    rq_activate_all_grippers(True)
    # end: URCap Program Node
  end
  $ 62 "zero_ftsensor()"
  zero_ftsensor()
  $ 63 "EXTT"
  $ 64 "Set GRP_3F_Enable=Off"
  set_standard_digital_out(4, False)
  $ 65 "Set BarcodeTrigger=Off"
  set_standard_digital_out(6, False)
  $ 66 "Set GRP_3F_Decap=Off"
  set_standard_digital_out(3, False)
  $ 67 "Set GRP_3F_Cap=Off"
  set_standard_digital_out(2, False)
  $ 68 "Set GRP_3F_Open=Off"
  set_standard_digital_out(5, False)
  $ 69 "PSE_T≔get_tool_free_pose(dir=[0,0,0.150], move_in_base_frame=True)"
  global PSE_T=get_tool_free_pose(dir=[0,0,0.150], move_in_base_frame=True)
  $ 70 "If is_reachable(Base_const, [PSE_T])"
  if (is_reachable(p[0.0,0.0,0.0,0.0,0.0,0.0], [PSE_T])):
    $ 71 "MoveL"
    $ 72 "PSE_T" "breakAfter"
    movel(PSE_T, a=1.2, v=0.15)
  end
  $ 74 "powder dispensing variable init"
  $ 75 "Start_thread≔ False "
  global Start_thread=  False
  $ 76 "vib_thread≔ False "
  global vib_thread=  False
  $ 77 "kp≔0.0015"
  global kp=0.0015
  $ 78 "ki≔0.0001"
  global ki=0.0001
  $ 79 "kd≔0.01"
  global kd=0.01
  $ 80 "dt≔0.03"
  global dt=0.03
  $ 81 "Integral_error≔0"
  global Integral_error=0
  $ 82 "current_error≔0"
  global current_error=0
  $ 83 "previous_error≔0"
  global previous_error=0
  $ 84 "tilt_increment≔0"
  global tilt_increment=0
  $ 85 "tilt_angle≔0"
  global tilt_angle=0
  $ 86 "diff≔0"
  global diff=0
  $ 87 "current_pose≔get_actual_tcp_pose()"
  global current_pose= get_actual_tcp_pose ()
  $ 88 "Relative_trans≔p[0, 0, -0.035, 0, 0, 0]"
  global Relative_trans=p[0, 0, -0.035, 0, 0, 0]
  $ 89 "ContA_plc_offst≔p[-0.00205, 0.02547, 0.03730, -0.03, -2.183, 6.165]"
  global ContA_plc_offst=p[-0.00205, 0.02547, 0.03730, -0.03, -2.183, 6.165]
  $ 90 "PowA_50_offset≔p[0.21808, -0.19943, 0.06584, 0, 0, 0]"
  global PowA_50_offset=p[0.21808, -0.19943, 0.06584, 0, 0, 0]
  $ 92 "tilt_init_reference()"
  tilt_init_reference()
  $ 93 "switch_spat_M≔ True "
  global switch_spat_M=  True
  $ 94 "switch_spat_S≔ True "
  global switch_spat_S=  True
  $ 95 "switch_spat_F_M≔ True "
  global switch_spat_F_M=  True
  $ 96 "switch_spat_F_S≔ True "
  global switch_spat_F_S=  True
  $ 97 "last_scale≔0"
  global last_scale=0
  $ 98 "W_EMPTY≔51.381"
  global W_EMPTY=51.381
  $ 771 "Thread_1"
  thread Thread_1():
    while (True):
      $ 772 "If Start_thread≟ True "
      if (Start_thread ==   True  ):
        $ 773 "weight_value≔get_weight()"
        global weight_value=get_weight()
        $ 774 "Wait: 0.1"
        sleep(0.1)
        $ 775 "sync()"
        sync()
      end
      $ 776 "sync()"
      sync()
    end
  end
  threadId_Thread_1 = run Thread_1()
  $ 777 "Thread_2"
  thread Thread_2():
    while (True):
      $ 778 "Loop vib_thread≟ True "
      thread Thread_while_778():
        while (True):
          $ 779 "diff≔target_weight-weight_value"
          global diff=target_weight-weight_value
          $ 780 "If diff>0.02 and spatula≠'spatula_flat_S'"
          global thread_flag_780=0
          thread Thread_if_780():
            $ 782 "Set AO[0]=4.0"
            set_standard_analog_out(0, 0.4)
            thread_flag_780 = 1
          end
          if (diff>0.02  and  spatula != "spatula_flat_S"):
            global thread_handler_780=run Thread_if_780()
            while (thread_flag_780 == 0):
              if not(diff>0.02  and  spatula != "spatula_flat_S"):
                kill thread_handler_780
                thread_flag_780 = 2
              else:
                sync()
              end
            end
          else:
            thread_flag_780 = 2
          end
          if (thread_flag_780 == 2):
            $ 783 "ElseIf diff>0.02 and spatula≟'spatula_flat_S'"
            if (diff>0.02 and spatula == "spatula_flat_S"):
              $ 784 "vibration_3()"
              vibration_3()
            else:
              $ 785 "ElseIf diff≤0.03"
              global thread_flag_785=0
              thread Thread_if_785():
                $ 786 "vibration_2()"
                vibration_2()
                thread_flag_785 = 1
              end
              if (diff <= 0.03):
                global thread_handler_785=run Thread_if_785()
                while (thread_flag_785 == 0):
                  if not(diff <= 0.03):
                    kill thread_handler_785
                    thread_flag_785 = 2
                  else:
                    sync()
                  end
                end
              else:
                thread_flag_785 = 2
              end
              if (thread_flag_785 == 2):
                $ 791 "Else" "noBreak"
                $ 792 "Set AO[0]=0.0"
                set_standard_analog_out(0, 0.0)
              end
            end
          end
        end
      end
      if (vib_thread ==   True  ):
        global thread_handler_778=run Thread_while_778()
        while (vib_thread ==   True  ):
          sync()
        end
        kill thread_handler_778
      end
      $ 793 "sync()"
      sync()
    end
  end
  threadId_Thread_2 = run Thread_2()
  while (True):
    $ 99 "Robot Program"
    $ 100 "MAIN"
    $ 101 "command_manager(external_control='uGO', cond_suspend=(ITM_Manipulated and AMR_AtTarget and AMR_Charging and AMR_Battery<40), cond_unsuspend=(AMR_Battery≟60))"
    command_manager(external_control="uGO", cond_suspend=(ITM_Manipulated  and  AMR_AtTarget  and  AMR_Charging  and  AMR_Battery<40), cond_unsuspend=(AMR_Battery == 60))
    $ 102 "log_state(STATE_Info)"
    log_state(STATE_Info)
    $ 103 "Switch STATE"
    switch_1 = STATE
    $ 104 "Case 1"
    if (1 == switch_1):
      $ 105 "Stopping"
      $ 106 "STATE_Info≔'Stopping'"
      global STATE_Info="Stopping"
      $ 107 "end_freedrive_mode()"
      end_freedrive_mode()
      $ 108 "Set"
      set_tcp(p[0.0,0.0,0.161,3.1415,0.0,0.0])
      $ 109 "PSE_T≔get_tool_free_pose(dir=[0,0,0.150], move_in_base_frame=True)"
      global PSE_T=get_tool_free_pose(dir=[0,0,0.150], move_in_base_frame=True)
      $ 110 "If is_reachable(Base_const, [PSE_T])"
      if (is_reachable(p[0.0,0.0,0.0,0.0,0.0,0.0], [PSE_T])):
        $ 111 "MoveL"
        $ 112 "PSE_T" "breakAfter"
        movel(PSE_T, a=1.2, v=0.15)
      end
      $ 113 "do_transition(keep_rxry=OBJ_Picked, r=0)"
      do_transition(keep_rxry=OBJ_Picked, r=0)
      $ 122 "Call Sub_AMR_MiR_V3"
      Sub_AMR_MiR_V3()
      $ 123 "If stopping() and AMR_Done"
      if (stopping()  and  AMR_Done):
        $ 124 "STATE≔2"
        global STATE=2
        $ 125 "ugo_update_outputs()"
        ugo_update_outputs()
      end
    elif (2 == switch_1):
      $ 126 "Case 2"
      $ 127 "Stopped"
      $ 128 "STATE_Info≔'Stopped'"
      global STATE_Info="Stopped"
      $ 129 "Call Sub_AMR_MiR_V3"
      Sub_AMR_MiR_V3()
      $ 130 "If CMD_Reset  or PB_Start"
      if (CMD_Reset   or  get_standard_digital_in(0)):
        $ 131 "STATE≔3"
        global STATE=3
        $ 132 "ugo_update_outputs()"
        ugo_update_outputs()
      end
    elif (3 == switch_1):
      $ 133 "Case 3"
      $ 134 " Resetting"
      $ 135 "STATE_Info≔'Resetting'"
      global STATE_Info="Resetting"
      $ 136 "uML"
      $ 137 "reset_error()"
      reset_error()
      $ 138 "reset_warning()"
      reset_warning()
      $ 139 "PROCESS_Step≔0"
      global PROCESS_Step=0
      $ 140 "PROCESS_Info≔''"
      global PROCESS_Info=""
      $ 141 "ARM_Referenced≔ False "
      global ARM_Referenced=  False
      $ 142 "WRK_Done≔ False "
      global WRK_Done=  False
      $ 143 "ITM_Prepared≔ False "
      global ITM_Prepared=  False
      $ 144 "ITM_Manipulated≔ False "
      global ITM_Manipulated=  False
      $ 145 "STP≔0"
      global STP=0
      $ 146 "Action≔0"
      global Action=0
      $ 147 "Action_Info≔''"
      global Action_Info=""
      $ 148 "ITM_ID≔0"
      global ITM_ID=0
      $ 149 "JIG≔0"
      global JIG=0
      $ 150 "JIG_Slot≔0"
      global JIG_Slot=0
      $ 151 "Task_info≔''"
      global Task_info=""
      $ 152 "Set"
      set_tcp(p[0.0,0.0,0.161,3.1415,0.0,0.0])
      $ 153 "App"
      $ 154 "'ADD APPLICATION SPECIFIC COMMANDS'"
      # 'ADD APPLICATION SPECIFIC COMMANDS'
      $ 155 "OBJ_Type≔0"
      global OBJ_Type=0
      $ 156 "OBJ_Nbr≔0"
      global OBJ_Nbr=0
      $ 157 "If CNT_Rack_Output≥50"
      if (CNT_Rack_Output >= 50):
        $ 158 "CNT_Rack_Output≔0"
        global CNT_Rack_Output=0
      end
      $ 159 "TASK≔struct(ID=0, NAVI=struct(target=0, footprint=0, protectiveOff=0, dock=0), WORK=struct(ITM_ID_Src=0, JIG_ID_Src=0, OBJ_Nbr_Src=0, ACT_Src=0, ITM_ID_Tgt=0, JIG_ID_Tgt=0, OBJ_Nbr_Tgt=0, ACT_Tgt=0, OBJ_Type=0))"
      global TASK=struct(ID=0, NAVI=struct(target=0, footprint=0, protectiveOff=0, dock=0), WORK=struct(ITM_ID_Src=0, JIG_ID_Src=0, OBJ_Nbr_Src=0, ACT_Src=0, ITM_ID_Tgt=0, JIG_ID_Tgt=0, OBJ_Nbr_Tgt=0, ACT_Tgt=0, OBJ_Type=0))
      $ 160 "Call Sub_AMR_MiR_V3"
      Sub_AMR_MiR_V3()
      $ 161 "If resetting() and AMR_Done"
      if (resetting()  and  AMR_Done):
        $ 162 "STATE≔4"
        global STATE=4
        $ 163 "ugo_update_outputs()"
        ugo_update_outputs()
      end
    elif (4 == switch_1):
      $ 164 "Case 4"
      $ 165 "Idle"
      $ 166 "STATE_Info≔'Idle'"
      global STATE_Info="Idle"
      $ 167 "If CMD_Start"
      if (CMD_Start):
        $ 168 "STATE≔5"
        global STATE=5
        $ 169 "ugo_update_outputs()"
        ugo_update_outputs()
      end
    elif (5 == switch_1):
      $ 170 "Case 5"
      $ 171 "Starting"
      $ 172 "STATE_Info≔'Starting'"
      global STATE_Info="Starting"
      $ 173 "'ADD COMMANDS WHAT TO START WITH'"
      # 'ADD COMMANDS WHAT TO START WITH'
      $ 174 "Call Sub_AMR_MiR_V3"
      Sub_AMR_MiR_V3()
      $ 175 "get ugo data"
      $ 176 "Assign Tasks"
      $ 177 "TASK.ID = ugo_get_task()"
      TASK.ID = ugo_get_task()
      $ 178 "If TASK.ID≟1"
      if (TASK.ID == 1):
        $ 179 "Task_info≔'Charge'"
        global Task_info="Charge"
        $ 180 "Parameters"
        $ 181 "AMR_PosTarget≔1"
        global AMR_PosTarget=1
      else:
        $ 182 "ElseIf TASK.ID≟9"
        if (TASK.ID == 9):
          $ 183 "'Pick Sarstedt Rack from Variable source'"
          # 'Pick Sarstedt Rack from Variable source'
          $ 184 "Task_info≔'Navigate to Target'"
          global Task_info="Navigate to Target"
          $ 185 "Parameters"
          $ 186 "AMR_PosTarget≔UGO.read_input('00','ITM_ID')"
          global AMR_PosTarget=UGO.read_input("00","ITM_ID")
        else:
          $ 187 "ElseIf TASK.ID≟49"
          if (TASK.ID == 49):
            $ 188 "Task_info≔'Pick Containers'"
            global Task_info="Pick Containers"
            $ 189 "Parameters"
            $ 190 "ITM_ID≔1"
            global ITM_ID=1
            $ 191 "OBJ_Type≔6"
            global OBJ_Type=6
            $ 192 "JIG≔15"
            global JIG=15
            $ 193 "AMR_PosTarget≔3"
            global AMR_PosTarget=3
          else:
            $ 194 "ElseIf TASK.ID≟50"
            if (TASK.ID == 50):
              $ 195 "Task_info≔'Decap Containers'"
              global Task_info="Decap Containers"
              $ 196 "Parameters"
              $ 197 "ITM_ID≔1"
              global ITM_ID=1
              $ 198 "OBJ_Type≔6"
              global OBJ_Type=6
              $ 199 "JIG≔16"
              global JIG=16
              $ 200 "AMR_PosTarget≔5"
              global AMR_PosTarget=5
            else:
              $ 201 "ElseIf TASK.ID≟51"
              if (TASK.ID == 51):
                $ 202 "Task_info≔'Detect Spatula and transfer powder'"
                global Task_info="Detect Spatula and transfer powder"
                $ 203 "Parameters"
                $ 204 "ITM_ID≔1"
                global ITM_ID=1
                $ 205 "target_weight≔(UGO.read_input('00','Target_weight'))/1000"
                global target_weight=(UGO.read_input("00","Target_weight"))/1000
                $ 206 "OBJ_Type≔8"
                global OBJ_Type=8
                $ 207 "JIG≔16"
                global JIG=16
                $ 208 "AMR_PosTarget≔5"
                global AMR_PosTarget=5
              else:
                $ 209 "ElseIf TASK.ID≟52"
                if (TASK.ID == 52):
                  $ 210 "Task_info≔'Pick Powder'"
                  global Task_info="Pick Powder"
                  $ 211 "Parameters"
                  $ 212 "ITM_ID≔1"
                  global ITM_ID=1
                  $ 213 "OBJ_Type≔6"
                  global OBJ_Type=6
                  $ 214 "JIG≔15"
                  global JIG=15
                  $ 215 "AMR_PosTarget≔3"
                  global AMR_PosTarget=3
                else:
                  $ 216 "ElseIf TASK.ID≟53"
                  if (TASK.ID == 53):
                    $ 217 "Task_info≔'Decap Powder'"
                    global Task_info="Decap Powder"
                    $ 218 "Parameters"
                    $ 219 "ITM_ID≔1"
                    global ITM_ID=1
                    $ 220 "OBJ_Type≔6"
                    global OBJ_Type=6
                    $ 221 "JIG≔1"
                    global JIG=1
                    $ 222 "AMR_PosTarget≔5"
                    global AMR_PosTarget=5
                  else:
                    $ 223 "ElseIf TASK.ID≟54"
                    if (TASK.ID == 54):
                      $ 224 "Task_info≔'Empty and swap Powder container'"
                      global Task_info="Empty and swap Powder container"
                      $ 233 "Parameters"
                      $ 234 "ITM_ID≔1"
                      global ITM_ID=1
                      $ 236 "W_now≔(UGO.read_input('00','Container_weight'))/1000"
                      global W_now=(UGO.read_input("00","Container_weight"))/1000
                      $ 237 "Pow_name≔(UGO.read_input('00','Powder_name'))"
                      global Pow_name=(UGO.read_input("00","Powder_name"))
                      $ 238 "scooping_init()"
                      scooping_init()
                      $ 239 "target_weight≔W_now-W_EMPTY-(0.002*W_FULL)"
                      global target_weight=W_now-W_EMPTY-(0.002*W_FULL)
                      $ 240 "OBJ_Type≔6"
                      global OBJ_Type=6
                      $ 241 "JIG≔17"
                      global JIG=17
                      $ 242 "AMR_PosTarget≔5"
                      global AMR_PosTarget=5
                    else:
                      $ 243 "ElseIf TASK.ID≟55"
                      if (TASK.ID == 55):
                        $ 244 "Task_info≔'Place Powder'"
                        global Task_info="Place Powder"
                        $ 245 "Parameters"
                        $ 246 "ITM_ID≔1"
                        global ITM_ID=1
                        $ 247 "OBJ_Type≔6"
                        global OBJ_Type=6
                        $ 248 "JIG≔21"
                        global JIG=21
                        $ 249 "AMR_PosTarget≔5"
                        global AMR_PosTarget=5
                      else:
                        $ 250 "ElseIf TASK.ID≟56"
                        if (TASK.ID == 56):
                          $ 251 "Task_info≔'Dose Powder'"
                          global Task_info="Dose Powder"
                          $ 252 "Parameters"
                          $ 253 "ITM_ID≔1"
                          global ITM_ID=1
                          $ 254 "target_weight≔(UGO.read_input('00','Target_weight'))/1000"
                          global target_weight=(UGO.read_input("00","Target_weight"))/1000
                          $ 255 "W_now≔(UGO.read_input('00','Container_weight'))/1000"
                          global W_now=(UGO.read_input("00","Container_weight"))/1000
                          $ 257 "Pow_name≔(UGO.read_input('00','Powder_name'))"
                          global Pow_name=(UGO.read_input("00","Powder_name"))
                          $ 258 "OBJ_Type≔6"
                          global OBJ_Type=6
                          $ 259 "JIG≔17"
                          global JIG=17
                          $ 260 "AMR_PosTarget≔5"
                          global AMR_PosTarget=5
                        else:
                          $ 261 "ElseIf TASK.ID≟57"
                          if (TASK.ID == 57):
                            $ 262 "Task_info≔'Recipe Powder dosing'"
                            global Task_info="Recipe Powder dosing"
                            $ 263 "Parameters"
                            $ 264 "ITM_ID≔1"
                            global ITM_ID=1
                            $ 265 "Pow_A≔(UGO.read_input('00','PowderA'))"
                            global Pow_A=(UGO.read_input("00","PowderA"))
                            $ 266 "Pow_B≔(UGO.read_input('00','PowderB'))"
                            global Pow_B=(UGO.read_input("00","PowderB"))
                            $ 267 "Pow_C≔(UGO.read_input('00','PowderC'))"
                            global Pow_C=(UGO.read_input("00","PowderC"))
                            $ 268 "Total_weight≔(UGO.read_input('00','Total_weight'))/1000"
                            global Total_weight=(UGO.read_input("00","Total_weight"))/1000
                            $ 269 "Pow_A_percent≔(UGO.read_input('00','PowderA_percentage'))/100"
                            global Pow_A_percent=(UGO.read_input("00","PowderA_percentage"))/100
                            $ 270 "Pow_B_percent≔(UGO.read_input('00','PowderB_percentage'))/100"
                            global Pow_B_percent=(UGO.read_input("00","PowderB_percentage"))/100
                            $ 271 "Pow_C_percent≔(UGO.read_input('00','PowderC_percentage'))/100"
                            global Pow_C_percent=(UGO.read_input("00","PowderC_percentage"))/100
                            $ 272 "OBJ_Type≔6"
                            global OBJ_Type=6
                            $ 273 "JIG≔17"
                            global JIG=17
                            $ 274 "AMR_PosTarget≔5"
                            global AMR_PosTarget=5
                          else:
                            $ 275 "ElseIf TASK.ID≟58"
                            if (TASK.ID == 58):
                              $ 276 "Task_info≔'Pick Powder containers'"
                              global Task_info="Pick Powder containers"
                              $ 277 "Parameters"
                              $ 278 "ITM_ID≔1"
                              global ITM_ID=1
                              $ 279 "OBJ_Type≔6"
                              global OBJ_Type=6
                              $ 280 "JIG≔15"
                              global JIG=15
                              $ 281 "AMR_PosTarget≔3"
                              global AMR_PosTarget=3
                            else:
                              $ 282 "Else" "noBreak"
                              $ 283 "set_error(ERROR_WRONG_ORDER)"
                              set_error(ERROR_WRONG_ORDER)
                            end
                          end
                        end
                      end
                    end
                  end
                end
              end
            end
          end
        end
      end
      $ 284 "test ugo"
      $ 285 "Wait: 0.2"
      sleep(0.2)
      $ 286 "ugo_update_outputs()"
      ugo_update_outputs()
      $ 287 "If starting() and AMR_Done"
      if (starting()  and  AMR_Done):
        $ 288 "log_message(Task_info, 'New Task: ')"
        log_message(Task_info, "New Task: ")
        $ 289 "log_message(to_str(TASK.ID), 'Task_ID: ')"
        log_message(to_str(TASK.ID), "Task_ID: ")
        $ 290 "do_transition(keep_rxry=OBJ_Picked)"
        do_transition(keep_rxry=OBJ_Picked)
        $ 291 "STATE≔6"
        global STATE=6
        $ 292 "ugo_update_outputs()"
        ugo_update_outputs()
      end
    elif (6 == switch_1):
      $ 293 "Case 6"
      $ 294 "Execute"
      $ 295 "STATE_Info≔'Execute'"
      global STATE_Info="Execute"
      $ 296 "If  not CMD_Hold and not CMD_Suspend"
      global thread_flag_296=0
      thread Thread_if_296():
        $ 297 "Switch PROCESS_Step"
        switch_2 = PROCESS_Step
        $ 298 "Case 0"
        if (0 == switch_2):
          $ 299 "PROCESS_Info≔'process control'"
          global PROCESS_Info="process control"
          $ 300 "log_process(PROCESS_Info)"
          log_process(PROCESS_Info)
          $ 301 "process control"
          $ 302 "If  not AMR_AtTarget"
          if (  not  AMR_AtTarget):
            $ 303 "PROCESS_Step≔1"
            global PROCESS_Step=1
          else:
            $ 304 "ElseIf (( not ITM_Prepared and  not WRK_Done) or (ITM_Prepared and WRK_Done))"
            if (((  not  ITM_Prepared  and    not  WRK_Done)  or  (ITM_Prepared  and  WRK_Done))):
              $ 305 "PROCESS_Step≔2"
              global PROCESS_Step=2
            else:
              $ 306 "ElseIf  not WRK_Done"
              if (  not  WRK_Done):
                $ 307 "PROCESS_Step≔3"
                global PROCESS_Step=3
              else:
                $ 308 "Else" "noBreak"
                $ 309 "task finished"
                $ 310 "PROCESS_Info≔''"
                global PROCESS_Info=""
                $ 311 "STATE≔7"
                global STATE=7
                $ 312 "ugo_update_outputs()"
                ugo_update_outputs()
              end
            end
          end
        elif (1 == switch_2):
          $ 313 "Case 1"
          $ 314 "navigate"
          $ 315 "'MOVING THE uML'"
          # 'MOVING THE uML'
          $ 316 "PROCESS_Info≔'move to target'"
          global PROCESS_Info="move to target"
          $ 317 "log_process(PROCESS_Info)"
          log_process(PROCESS_Info)
          $ 318 "If TASK.ID≟1"
          if (TASK.ID == 1):
            $ 319 "Action≔51"
            global Action=51
          else:
            $ 320 "Else" "noBreak"
            $ 321 "Action≔52"
            global Action=52
          end
          $ 322 "Call Sub_AMR_MiR_V3"
          Sub_AMR_MiR_V3()
          $ 323 "If AMR_Done"
          if (AMR_Done):
            $ 324 "PROCESS_Step≔0"
            global PROCESS_Step=0
          end
        elif (2 == switch_2):
          $ 325 "Case 2"
          $ 326 "prepare"
          $ 327 "'THINGS THAT HAVE TO BE DONE ONCE IN A SEQUENCE,WORKFLOW'"
          # 'THINGS THAT HAVE TO BE DONE ONCE IN A SEQUENCE,WORKFLOW'
          $ 328 "PROCESS_Info≔'prepare for work'"
          global PROCESS_Info="prepare for work"
          $ 329 "log_process(PROCESS_Info)"
          log_process(PROCESS_Info)
          $ 330 "If TASK.WORK.ITM_ID_Src>1"
          if (TASK.WORK.ITM_ID_Src>1):
            $ 331 "ITM_ID≔TASK.WORK.ITM_ID_Src"
            global ITM_ID=TASK.WORK.ITM_ID_Src
          else:
            $ 332 "ElseIf TASK.WORK.ITM_ID_Tgt>1"
            if (TASK.WORK.ITM_ID_Tgt>1):
              $ 333 "ITM_ID≔TASK.WORK.ITM_ID_Tgt"
              global ITM_ID=TASK.WORK.ITM_ID_Tgt
            end
          end
          $ 334 "If  not ARM_Referenced and (ITM_ID≠0)"
          if (  not  ARM_Referenced  and  (ITM_ID != 0)):
            $ 335 "STP≔1"
            global STP=1
          else:
            $ 336 "ElseIf ARM_Referenced or (ITM_ID≟0)"
            if (ARM_Referenced  or  (ITM_ID == 0)):
              $ 337 "STP≔2"
              global STP=2
            end
          end
          $ 338 "Switch STP"
          switch_3 = STP
          $ 339 "Case 1"
          if (1 == switch_3):
            $ 340 "reference"
            $ 341 "STP_Info≔'reference at target position'"
            global STP_Info="reference at target position"
            $ 342 "log_step(STP_Info)"
            log_step(STP_Info)
            $ 343 "If ITM_ID≟1"
            if (ITM_ID == 1):
              $ 344 "CAM_Done≔ True "
              global CAM_Done=  True
            else:
              $ 345 "Else" "noBreak"
              $ 346 "Action≔131"
              global Action=131
              $ 347 "Call Sub_Vision_V18"
              Sub_Vision_V18()
            end
            $ 349 "If CAM_Done and  not ERROR.FLAG"
            if (CAM_Done  and    not  ERROR.FLAG):
              $ 350 "log_step('ARM referenced')"
              log_step("ARM referenced")
              $ 351 "ARM_Referenced≔ True "
              global ARM_Referenced=  True
            end
          elif (2 == switch_3):
            $ 352 "Case 2"
            $ 353 "manipulate"
            $ 354 "STP_Info≔'manipulate item'"
            global STP_Info="manipulate item"
            $ 355 "log_step(STP_Info)"
            log_step(STP_Info)
            $ 356 "'In case pressing button is needed'"
            # 'In case pressing button is needed'
            $ 357 "If found_in_list(ITM_ID, ITM_ID_List)"
            if (found_in_list(ITM_ID, ITM_ID_List)):
              $ 358 "Switch ITM_ID"
              switch_4 = ITM_ID
              $ 359 "Case 0"
              if (0 == switch_4):
                $ 360 "ITM_Manipulated≔ not ITM_Manipulated"
                global ITM_Manipulated=  not  ITM_Manipulated
              elif (1 == switch_4):
                $ 361 "Case 1"
                $ 362 "ITM_Manipulated≔ not ITM_Manipulated"
                global ITM_Manipulated=  not  ITM_Manipulated
              elif (2 == switch_4):
                $ 363 "Case 2"
              else:
                $ 373 "Default Case"
                $ 374 "ITM_Manipulated≔ not ITM_Manipulated"
                global ITM_Manipulated=  not  ITM_Manipulated
              end
            end
          end
          $ 375 "ITM_Prepared≔(ITM_Manipulated or  not found_in_list(ITM_ID, ITM_ID_List)) and (ARM_Referenced or ITM_ID≟0) and  not WRK_Done"
          global ITM_Prepared=(ITM_Manipulated  or    not  found_in_list(ITM_ID, ITM_ID_List))  and  (ARM_Referenced  or  ITM_ID == 0)  and    not  WRK_Done
          $ 376 "STP≔0"
          global STP=0
          $ 377 "STP_Info≔''"
          global STP_Info=""
          $ 378 "PROCESS_Step≔0"
          global PROCESS_Step=0
        elif (3 == switch_2):
          $ 379 "Case 3"
          $ 380 "work"
          $ 381 "'ADD EVERY MACHINE, OBJECT, STATION TO WORK ON'"
          # 'ADD EVERY MACHINE, OBJECT, STATION TO WORK ON'
          $ 382 "Switch ITM_ID"
          switch_3 = ITM_ID
          $ 383 "Case 1"
          if (1 == switch_3):
            $ 384 "uLM"
            $ 385 "If TASK.ID≟12"
            if (TASK.ID == 12):
              $ 386 "fill racks"
              $ 387 "Action≔151"
              global Action=151
              $ 388 "Call Sub_Vision_V18"
              Sub_Vision_V18()
              $ 389 "If  not ERROR.FLAG"
              if (  not  ERROR.FLAG):
                $ 390 "Actions for the task"
                $ 391 "Action≔1"
                global Action=1
                $ 392 "JIG≔2"
                global JIG=2
                $ 393 "JIG_Slot≔CAM_Result[0]"
                global JIG_Slot=CAM_Result[0]
                $ 394 "OBJ_Nbr≔CAM_Result[0]"
                global OBJ_Nbr=CAM_Result[0]
                $ 395 "OBJ_Type≔2"
                global OBJ_Type=2
                $ 396 "Call Sub_Action_V4"
                Sub_Action_V4()
                $ 397 "If OBJ_Picked"
                if (OBJ_Picked):
                  $ 398 "CAM_Result.remove(0)"
                  CAM_Result.remove(0)
                  $ 399 "PRC_TubCounter≔PRC_TubCounter+1"
                  global PRC_TubCounter=PRC_TubCounter+1
                  $ 400 "If PRC_TubCounter%4≟0"
                  if (PRC_TubCounter%4 == 0):
                    $ 401 "JIG_Slot≔4"
                    global JIG_Slot=4
                  else:
                    $ 402 "Else" "noBreak"
                    $ 403 "JIG_Slot≔PRC_TubCounter%4"
                    global JIG_Slot=PRC_TubCounter%4
                  end
                  $ 404 "OBJ_Nbr≔ceil(PRC_TubCounter/4)"
                  global OBJ_Nbr=ceil(PRC_TubCounter/4)
                  $ 405 "Action≔2"
                  global Action=2
                  $ 406 "JIG≔4"
                  global JIG=4
                  $ 407 "Call Sub_Action_V4"
                  Sub_Action_V4()
                  $ 408 "Action≔151"
                  global Action=151
                  $ 409 "Call Sub_Vision_V18"
                  Sub_Vision_V18()
                end
              end
              $ 410 "If (CAM_Captures≥CAM_PRM_Retries) or (PRC_TubCounter≥32)"
              if ((CAM_Captures >= CAM_PRM_Retries)  or  (PRC_TubCounter >= 32)):
                $ 411 "PROCESS_Step≔0"
                global PROCESS_Step=0
                $ 412 "WRK_Done≔ True "
                global WRK_Done=  True
              end
            else:
              $ 413 "ElseIf TASK.ID≟49"
              if (TASK.ID == 49):
                $ 414 "Pick Powder container"
                $ 415 "Action≔131"
                global Action=131
                $ 416 "Call Sub_Vision_V18"
                Sub_Vision_V18()
                $ 417 "Action≔35"
                global Action=35
                $ 418 "Call Sub_Action_V4"
                Sub_Action_V4()
                $ 419 "PROCESS_Step≔0"
                global PROCESS_Step=0
                $ 420 "WRK_Done≔ True "
                global WRK_Done=  True
              else:
                $ 421 "ElseIf TASK.ID≟50"
                if (TASK.ID == 50):
                  $ 422 "Decap containers"
                  $ 423 "Action≔36"
                  global Action=36
                  $ 424 "Call Sub_Action_V4"
                  Sub_Action_V4()
                  $ 425 "PROCESS_Step≔0"
                  global PROCESS_Step=0
                  $ 426 "WRK_Done≔ True "
                  global WRK_Done=  True
                else:
                  $ 427 "ElseIf TASK.ID≟51"
                  if (TASK.ID == 51):
                    $ 428 "Detect Spatula and transfer powder"
                    $ 429 "Action≔131"
                    global Action=131
                    $ 430 "Call Sub_Vision_V18"
                    Sub_Vision_V18()
                    $ 431 "Action≔37"
                    global Action=37
                    $ 432 "Call Sub_Action_V4"
                    Sub_Action_V4()
                    $ 433 "PROCESS_Step≔0"
                    global PROCESS_Step=0
                    $ 434 "WRK_Done≔ True "
                    global WRK_Done=  True
                  else:
                    $ 435 "ElseIf TASK.ID≟52"
                    if (TASK.ID == 52):
                      $ 436 "Pick Powder container"
                      $ 437 "Action≔131"
                      global Action=131
                      $ 438 "Call Sub_Vision_V18"
                      Sub_Vision_V18()
                      $ 439 "Action≔39"
                      global Action=39
                      $ 440 "Call Sub_Action_V4"
                      Sub_Action_V4()
                      $ 441 "PROCESS_Step≔0"
                      global PROCESS_Step=0
                      $ 442 "WRK_Done≔ True "
                      global WRK_Done=  True
                    else:
                      $ 443 "ElseIf TASK.ID≟53"
                      if (TASK.ID == 53):
                        $ 444 "Decap containerA"
                        $ 445 "Action≔40"
                        global Action=40
                        $ 446 "Call Sub_Action_V4"
                        Sub_Action_V4()
                        $ 447 "PROCESS_Step≔0"
                        global PROCESS_Step=0
                        $ 448 "WRK_Done≔ True "
                        global WRK_Done=  True
                      else:
                        $ 449 "ElseIf TASK.ID≟55"
                        if (TASK.ID == 55):
                          $ 450 "Place Powder"
                          $ 451 "Action≔131"
                          global Action=131
                          $ 452 "Call Sub_Vision_V18"
                          Sub_Vision_V18()
                          $ 453 "Action≔41"
                          global Action=41
                          $ 454 "Call Sub_Action_V4"
                          Sub_Action_V4()
                          $ 455 "PROCESS_Step≔0"
                          global PROCESS_Step=0
                          $ 456 "WRK_Done≔ True "
                          global WRK_Done=  True
                        else:
                          $ 457 "ElseIf TASK.ID≟54"
                          if (TASK.ID == 54):
                            $ 458 "Empty and swap container"
                            $ 459 "Action≔131"
                            global Action=131
                            $ 460 "Call Sub_Vision_V18"
                            Sub_Vision_V18()
                            $ 461 "Action≔42"
                            global Action=42
                            $ 462 "Call Sub_Action_V4"
                            Sub_Action_V4()
                            $ 463 "PROCESS_Step≔0"
                            global PROCESS_Step=0
                            $ 464 "WRK_Done≔ True "
                            global WRK_Done=  True
                          else:
                            $ 465 "ElseIf TASK.ID≟56"
                            if (TASK.ID == 56):
                              $ 466 "Dispense Powder"
                              $ 467 "Action≔131"
                              global Action=131
                              $ 468 "Call Sub_Vision_V18"
                              Sub_Vision_V18()
                              $ 469 "Action≔43"
                              global Action=43
                              $ 470 "Call Sub_Action_V4"
                              Sub_Action_V4()
                              $ 471 "PROCESS_Step≔0"
                              global PROCESS_Step=0
                              $ 472 "WRK_Done≔ True "
                              global WRK_Done=  True
                            else:
                              $ 473 "ElseIf TASK.ID≟57"
                              if (TASK.ID == 57):
                                $ 474 "Recipe Dosing"
                                $ 475 "Action≔48"
                                global Action=48
                                $ 476 "Call Sub_Action_V4"
                                Sub_Action_V4()
                                $ 477 "recipe_init(Pow_A, Pow_B, Pow_C, Total_weight, Pow_A_percent, Pow_B_percent, Pow_C_percent)"
                                recipe_init(Pow_A, Pow_B, Pow_C, Total_weight, Pow_A_percent, Pow_B_percent, Pow_C_percent)
                                $ 478 "Loop recipe_next()≟ True "
                                while (recipe_next() ==   True  ):
                                  $ 479 "Action≔44"
                                  global Action=44
                                  $ 480 "Call Sub_Action_V4"
                                  Sub_Action_V4()
                                  $ 481 "JIG≔21"
                                  global JIG=21
                                  $ 482 "Action≔131"
                                  global Action=131
                                  $ 483 "Call Sub_Vision_V18"
                                  Sub_Vision_V18()
                                  $ 484 "Action≔45"
                                  global Action=45
                                  $ 485 "Call Sub_Action_V4"
                                  Sub_Action_V4()
                                  $ 486 "dosing_start()"
                                  dosing_start()
                                  $ 487 "JIG≔17"
                                  global JIG=17
                                  $ 488 "Action≔131"
                                  global Action=131
                                  $ 489 "Call Sub_Vision_V18"
                                  Sub_Vision_V18()
                                  $ 490 "Action≔46"
                                  global Action=46
                                  $ 491 "Call Sub_Action_V4"
                                  Sub_Action_V4()
                                  $ 492 "dosing_end()"
                                  dosing_end()
                                end
                                $ 493 "PROCESS_Step≔0"
                                global PROCESS_Step=0
                                $ 494 "WRK_Done≔ True "
                                global WRK_Done=  True
                              else:
                                $ 495 "ElseIf TASK.ID≟58"
                                if (TASK.ID == 58):
                                  $ 496 "Pick Powder containers"
                                  $ 497 "Num_cont_picked≔0"
                                  global Num_cont_picked=0
                                  $ 498 "powder_position≔'Position1'"
                                  global powder_position="Position1"
                                  $ 499 "Loop Num_cont_picked<3"
                                  while (Num_cont_picked<3):
                                    $ 500 "Action≔131"
                                    global Action=131
                                    $ 501 "Call Sub_Vision_V18"
                                    Sub_Vision_V18()
                                    $ 502 "Action≔47"
                                    global Action=47
                                    $ 503 "Call Sub_Action_V4"
                                    Sub_Action_V4()
                                  end
                                  $ 504 "PROCESS_Step≔0"
                                  global PROCESS_Step=0
                                  $ 505 "WRK_Done≔ True "
                                  global WRK_Done=  True
                                end
                              end
                            end
                          end
                        end
                      end
                    end
                  end
                end
              end
            end
          elif (2 == switch_3):
            $ 506 "Case 2"
          elif (5 == switch_3):
            $ 548 "Case 5"
          elif (20 == switch_3):
            $ 556 "Case 20"
          elif (43 == switch_3):
            $ 618 "Case 43"
          else:
            $ 626 "Default Case"
            $ 627 "WRK_Done≔ True "
            global WRK_Done=  True
            $ 628 "PROCESS_Step≔0"
            global PROCESS_Step=0
          end
        end
        thread_flag_296 = 1
      end
      if (  not  CMD_Hold and not CMD_Suspend):
        global thread_handler_296=run Thread_if_296()
        while (thread_flag_296 == 0):
          if not(  not  CMD_Hold and not CMD_Suspend):
            kill thread_handler_296
            thread_flag_296 = 2
          else:
            sync()
          end
        end
      else:
        thread_flag_296 = 2
      end
      $ 629 "If CMD_Hold"
      if (CMD_Hold):
        $ 630 "STATE≔9"
        global STATE=9
        $ 631 "ugo_update_outputs()"
        ugo_update_outputs()
      else:
        $ 632 "ElseIf CMD_Suspend"
        if (CMD_Suspend):
          $ 633 "STATE≔12"
          global STATE=12
          $ 634 "ugo_update_outputs()"
          ugo_update_outputs()
        end
      end
    elif (7 == switch_1):
      $ 635 "Case 7"
      $ 636 "Completing"
      $ 637 "STATE_Info≔'Completing'"
      global STATE_Info="Completing"
      $ 638 "'ADD COMMANDS FOR COMPLETING THE PROCESS'"
      # 'ADD COMMANDS FOR COMPLETING THE PROCESS'
      $ 639 "do_transition(keep_rxry=OBJ_Picked)"
      do_transition(keep_rxry=OBJ_Picked)
      $ 640 "Call Sub_AMR_MiR_V3"
      Sub_AMR_MiR_V3()
      $ 641 "If completing() and AMR_Done"
      if (completing()  and  AMR_Done):
        $ 642 "STATE≔8"
        global STATE=8
        $ 643 "ugo_update_outputs()"
        ugo_update_outputs()
      end
    elif (8 == switch_1):
      $ 644 "Case 8"
      $ 645 "Complete"
      $ 646 "STATE_Info≔'Complete'"
      global STATE_Info="Complete"
      $ 647 "If CMD_Reset"
      if (CMD_Reset):
        $ 648 "STATE≔3"
        global STATE=3
        $ 649 "ugo_update_outputs()"
        ugo_update_outputs()
      end
    elif (9 == switch_1):
      $ 650 "Case 9"
      $ 651 "Holding"
      $ 652 "STATE_Info≔'Holding'"
      global STATE_Info="Holding"
      $ 653 "stopl(0.5)"
      stopl(0.5)
      $ 654 "Call Sub_AMR_MiR_V3"
      Sub_AMR_MiR_V3()
      $ 655 "If holding() and AMR_Done"
      if (holding()  and  AMR_Done):
        $ 656 "STATE≔10"
        global STATE=10
        $ 657 "ugo_update_outputs()"
        ugo_update_outputs()
      end
    elif (10 == switch_1):
      $ 658 "Case 10"
      $ 659 "Held"
      $ 660 "STATE_Info≔'Held'"
      global STATE_Info="Held"
      $ 661 "If CMD_Unhold"
      if (CMD_Unhold):
        $ 662 "end_freedrive_mode()"
        end_freedrive_mode()
        $ 663 "STATE≔11"
        global STATE=11
        $ 664 "ugo_update_outputs()"
        ugo_update_outputs()
      else:
        $ 665 "ElseIf FNC_Freedrive"
        if (FNC_Freedrive):
          $ 666 "freedrive_mode()"
          freedrive_mode()
        else:
          $ 667 "Else" "noBreak"
          $ 668 "end_freedrive_mode()"
          end_freedrive_mode()
        end
      end
    elif (11 == switch_1):
      $ 669 "Case 11"
      $ 670 "Unholding"
      $ 671 "STATE_Info≔'Unholding'"
      global STATE_Info="Unholding"
      $ 672 "Clearing"
      $ 673 "Switch ERROR.ID"
      switch_2 = ERROR.ID
      $ 674 "Case 1002"
      if (1002 == switch_2):
        $ 675 "AMR_AtTarget≔ False "
        global AMR_AtTarget=  False
        $ 676 "ARM_Referenced≔ False "
        global ARM_Referenced=  False
        $ 677 "ITM_Prepared≔ False "
        global ITM_Prepared=  False
        $ 678 "PROCESS_Step≔1"
        global PROCESS_Step=1
      elif (2007 == switch_2):
        $ 679 "Case 2007"
        $ 680 "PROCESS_Step≔1"
        global PROCESS_Step=1
      end
      $ 681 "reset_error()"
      reset_error()
      $ 682 "reset_warning()"
      reset_warning()
      $ 683 "OBJ_Picked≔gripper_has_object()"
      global OBJ_Picked=gripper_has_object()
      $ 684 "Call Sub_AMR_MiR_V3"
      Sub_AMR_MiR_V3()
      $ 685 "If unholding() and AMR_Done"
      if (unholding()  and  AMR_Done):
        $ 686 "STATE≔6"
        global STATE=6
        $ 687 "ugo_update_outputs()"
        ugo_update_outputs()
      end
    elif (12 == switch_1):
      $ 688 "Case 12"
      $ 689 "Suspending"
      $ 690 "STATE_Info≔'Suspending'"
      global STATE_Info="Suspending"
      $ 691 "PROCESS_Info≔str_cat(PROCESS_Info, ' suspended')"
      global PROCESS_Info=str_cat(PROCESS_Info, " suspended")
      $ 692 "If suspending()"
      if (suspending()):
        $ 693 "STATE≔13"
        global STATE=13
        $ 694 "ugo_update_outputs()"
        ugo_update_outputs()
      end
    elif (13 == switch_1):
      $ 695 "Case 13"
      $ 696 "Suspended"
      $ 697 "STATE_Info≔'Suspended'"
      global STATE_Info="Suspended"
      $ 698 "Call Sub_AMR_MiR_V3"
      Sub_AMR_MiR_V3()
      $ 699 "If CMD_Unsuspend"
      if (CMD_Unsuspend):
        $ 700 "STATE≔14"
        global STATE=14
        $ 701 "ugo_update_outputs()"
        ugo_update_outputs()
      end
    elif (14 == switch_1):
      $ 702 "Case 14"
      $ 703 "Unsuspending"
      $ 704 "STATE_Info≔'Unsuspending'"
      global STATE_Info="Unsuspending"
      $ 705 "PROCESS_Step≔0"
      global PROCESS_Step=0
      $ 706 "If unsuspending()"
      if (unsuspending()):
        $ 707 "STATE≔6"
        global STATE=6
        $ 708 "ugo_update_outputs()"
        ugo_update_outputs()
      end
    elif (15 == switch_1):
      $ 709 "Case 15"
      $ 710 "Aborting"
      $ 711 "STATE_Info≔'Aborting'"
      global STATE_Info="Aborting"
      $ 712 "If aborting()"
      if (aborting()):
        $ 713 "STATE≔16"
        global STATE=16
        $ 714 "ugo_update_outputs()"
        ugo_update_outputs()
      end
    elif (16 == switch_1):
      $ 715 "Case 16"
      $ 716 "Aborted"
      $ 717 "STATE_Info≔'Aborted'"
      global STATE_Info="Aborted"
      $ 718 "If CMD_Clear"
      if (CMD_Clear):
        $ 719 "STATE≔17"
        global STATE=17
        $ 720 "ugo_update_outputs()"
        ugo_update_outputs()
      end
    elif (17 == switch_1):
      $ 721 "Case 17"
      $ 722 "Clearing"
      $ 723 "STATE_Info≔'Clearing'"
      global STATE_Info="Clearing"
      $ 724 "Clearing"
      $ 725 "reset_warning()"
      reset_warning()
      $ 726 "reset_error()"
      reset_error()
      $ 727 "If clearing()"
      if (clearing()):
        $ 728 "STATE≔2"
        global STATE=2
        $ 729 "ugo_update_outputs()"
        ugo_update_outputs()
      end
    end
    $ 730 "log_state(STATE_Info)"
    log_state(STATE_Info)
    $ 731 "log_warning(WARNING.MSG)"
    log_warning(WARNING.MSG)
    $ 732 "log_error(ERROR.MSG)"
    log_error(ERROR.MSG)
    $ 733 "Times"
    $ 734 "Switch STATE"
    switch_1 = STATE
    $ 735 "Case 1"
    if (1 == switch_1):
      $ 736 "TM_St_Stopping≔get_time(STATE_Times[STATE-1])"
      global TM_St_Stopping=get_time(STATE_Times[STATE-1])
    elif (2 == switch_1):
      $ 737 "Case 2"
      $ 738 "TM_St_Stopped≔get_time(STATE_Times[STATE-1])"
      global TM_St_Stopped=get_time(STATE_Times[STATE-1])
    elif (3 == switch_1):
      $ 739 "Case 3"
      $ 740 "TM_St_Resetting≔get_time(STATE_Times[STATE-1])"
      global TM_St_Resetting=get_time(STATE_Times[STATE-1])
    elif (4 == switch_1):
      $ 741 "Case 4"
      $ 742 "TM_St_Idle≔get_time(STATE_Times[STATE-1])"
      global TM_St_Idle=get_time(STATE_Times[STATE-1])
    elif (5 == switch_1):
      $ 743 "Case 5"
      $ 744 "TM_St_Starting≔get_time(STATE_Times[STATE-1])"
      global TM_St_Starting=get_time(STATE_Times[STATE-1])
    elif (6 == switch_1):
      $ 745 "Case 6"
      $ 746 "TM_St_Execute≔get_time(STATE_Times[STATE-1])"
      global TM_St_Execute=get_time(STATE_Times[STATE-1])
    elif (7 == switch_1):
      $ 747 "Case 7"
      $ 748 "TM_St_Completin≔get_time(STATE_Times[STATE-1])"
      global TM_St_Completin=get_time(STATE_Times[STATE-1])
    elif (8 == switch_1):
      $ 749 "Case 8"
      $ 750 "TM_St_Complete≔get_time(STATE_Times[STATE-1])"
      global TM_St_Complete=get_time(STATE_Times[STATE-1])
    elif (9 == switch_1):
      $ 751 "Case 9"
      $ 752 "TM_St_Holding≔get_time(STATE_Times[STATE-1])"
      global TM_St_Holding=get_time(STATE_Times[STATE-1])
    elif (10 == switch_1):
      $ 753 "Case 10"
      $ 754 "TM_St_Held≔get_time(STATE_Times[STATE-1])"
      global TM_St_Held=get_time(STATE_Times[STATE-1])
    elif (11 == switch_1):
      $ 755 "Case 11"
      $ 756 "TM_St_Unholding≔get_time(STATE_Times[STATE-1])"
      global TM_St_Unholding=get_time(STATE_Times[STATE-1])
    elif (12 == switch_1):
      $ 757 "Case 12"
      $ 758 "TM_St_Suspendin≔get_time(STATE_Times[STATE-1])"
      global TM_St_Suspendin=get_time(STATE_Times[STATE-1])
    elif (13 == switch_1):
      $ 759 "Case 13"
      $ 760 "TM_St_Suspended≔get_time(STATE_Times[STATE-1])"
      global TM_St_Suspended=get_time(STATE_Times[STATE-1])
    elif (14 == switch_1):
      $ 761 "Case 14"
      $ 762 "TM_St_Unsuspend≔get_time(STATE_Times[STATE-1])"
      global TM_St_Unsuspend=get_time(STATE_Times[STATE-1])
    elif (15 == switch_1):
      $ 763 "Case 15"
      $ 764 "TM_St_Aborting≔get_time(STATE_Times[STATE-1])"
      global TM_St_Aborting=get_time(STATE_Times[STATE-1])
    elif (16 == switch_1):
      $ 765 "Case 16"
      $ 766 "TM_St_Aborted≔get_time(STATE_Times[STATE-1])"
      global TM_St_Aborted=get_time(STATE_Times[STATE-1])
    elif (17 == switch_1):
      $ 767 "Case 17"
      $ 768 "TM_St_Clearing≔get_time(STATE_Times[STATE-1])"
      global TM_St_Clearing=get_time(STATE_Times[STATE-1])
    end
    $ 770 "Wait: 0.1"
    sleep(0.1)
  end
end
